ABB RAPID module: Module1.mod

MODULE Module1
	TASK PERS tooldata swieczka:=[TRUE,[[-64.6298,0.0716233,289.296],[1,0,0,0]],[1,[0,0,0],[1,0,0,0],0,0,0]];
    !***********************************************************
    !
    ! Module:  Module1
    !
    ! Description:
    !   <Insert description here>
    !
    ! Author: Mirgi
    !
    ! Version: 1.0
    !
    !***********************************************************


    !***********************************************************
    !
    ! Procedure main
    !
    !   This is the entry point of your program
    !
    !***********************************************************
    PROC main()
        !Add your code here
    ENDPROC
ENDMODULE
